Fanuc KAREL source: KT00807.KL

PROGRAM KT00807
%NOLOCKGROUP
VAR
  S1: STRING[80]
  S2: STRING[80]
  OUT: REAL
BEGIN
  S1 = 'A'
  S2 = 'B'
  S1 = 'A'
  S2 = 'B'
  OUT = EXP(S1)
END KT00807
